# EPICS substitutions: db/Beckhoff_5XXX/ecmcEL5101-0011.substitutions
file "ecmcEL5101-0011-chX.template"
{
  pattern { CH_ID, DTYP,             FTVL }
          { 01,    asynInt32ArrayIn, LONG }
}

# timestamp
file "ecmc_timestamp_64-chX.template"{
  pattern {CH_ID, KEY,      suffix,        sourceName         }
          {"",    "Enc01",   "-Time",       "nextSyncTime"    }
}
